(* IEC 61131-3 sources: 2026_Projet_YGO_ExcavatriceDragage/TOOLS/TEST_AUTO_CI/RESULTS/I_TRANSLATION/reports (part 3) *)

    ASSERT_FALSE(RestartSeen, 'aucun front montant mot/frequence apres l armement du verrou');
    ASSERT_TRUE(FB_T.ArrivalStopConfirmed, 'l arret confirme resiste au rebond et a la re-demande');
END_TEST

TEST 'TC-P11-037 T345-L1 Le fait d arret confirme n est ni constant ni efface par la demande'
    CfgFast.CfgRampAccelRate := 1000.0;
    CfgFast.CfgRampDecelNormalRate := 1000.0;
    CfgFast.CaptorDebounce := T#100ms;
    CfgFast.BrakeDelayMagnetise := T#0ms;
    CfgFast.BrakeDelayContactClose := T#0ms;

    (* Scan 1 : au repos, aucun arret confirme (le fait n est pas constant) *)
    FB_T(Enable := TRUE, Reset := FALSE, RunRequest := FALSE, SafeStop := FALSE,
         ReqTremie := FALSE, ReqMaintenance := FALSE, SpeedTgt_Pct := 50.0,
         PowerContactorEngaged := TRUE, Cfg := CfgFast,
         BypassContactorCheck := TRUE, BrakeFeedback := TRUE);
    ASSERT_FALSE(FB_T.ArrivalStopConfirmed, 'au repos : aucun arret confirme (fait non constant)');
    ADVANCE_TIME(10000000);

    (* Scans 2-5 : mouvement vers la cible *)
    FB_T(Enable := TRUE, Reset := FALSE, RunRequest := TRUE, SafeStop := FALSE,
         ReqTremie := TRUE, ReqMaintenance := FALSE, EffectivePermitM3_Tremie := TRUE,
         SpeedTgt_Pct := 50.0, PowerContactorEngaged := TRUE, Cfg := CfgFast,
         BypassContactorCheck := TRUE, BrakeFeedback := TRUE);
    ADVANCE_TIME(10000000);
    FB_T(Enable := TRUE, Reset := FALSE, RunRequest := TRUE, SafeStop := FALSE,
         ReqTremie := TRUE, ReqMaintenance := FALSE, EffectivePermitM3_Tremie := TRUE,
         SpeedTgt_Pct := 50.0, PowerContactorEngaged := TRUE, Cfg := CfgFast,
         BypassContactorCheck := TRUE, BrakeFeedback := TRUE);
    ADVANCE_TIME(10000000);
    FB_T(Enable := TRUE, Reset := FALSE, RunRequest := TRUE, SafeStop := FALSE,
         ReqTremie := TRUE, ReqMaintenance := FALSE, EffectivePermitM3_Tremie := TRUE,
         SpeedTgt_Pct := 50.0, PowerContactorEngaged := TRUE, Cfg := CfgFast,
         BypassContactorCheck := TRUE, BrakeFeedback := TRUE);
    ADVANCE_TIME(10000000);
    FB_T(Enable := TRUE, Reset := FALSE, RunRequest := TRUE, SafeStop := FALSE,
         ReqTremie := TRUE, ReqMaintenance := FALSE, EffectivePermitM3_Tremie := TRUE,
         SpeedTgt_Pct := 50.0, PowerContactorEngaged := TRUE, Cfg := CfgFast,
         BypassContactorCheck := TRUE, BrakeFeedback := TRUE);
    ASSERT_FALSE(FB_T.ArrivalStopConfirmed, 'en mouvement : aucun arret confirme');
    ADVANCE_TIME(10000000);

    (* Scans 6-20 : capteur cible, puis demande retiree avant la fin du debounce *)
    FB_T(Enable := TRUE, Reset := FALSE, RunRequest := TRUE, SafeStop := FALSE,
         ReqTremie := TRUE, ReqMaintenance := FALSE, EffectivePermitM3_Tremie := TRUE,
         SpeedTgt_Pct := 50.0, PowerContactorEngaged := TRUE, PositionSensorTarget := TRUE,
         Cfg := CfgFast, BypassContactorCheck := TRUE, BrakeFeedback := TRUE);
    ADVANCE_TIME(10000000);
    FB_T(Enable := TRUE, Reset := FALSE, RunRequest := FALSE, SafeStop := FALSE,
         ReqTremie := FALSE, ReqMaintenance := FALSE, EffectivePermitM3_Tremie := TRUE,
         SpeedTgt_Pct := 50.0, PowerContactorEngaged := TRUE, PositionSensorTarget := TRUE,
         Cfg := CfgFast, BypassContactorCheck := TRUE, BrakeFeedback := TRUE);
    ADVANCE_TIME(10000000);
    FB_T(Enable := TRUE, Reset := FALSE, RunRequest := FALSE, SafeStop := FALSE,
         ReqTremie := FALSE, ReqMaintenance := FALSE, EffectivePermitM3_Tremie := TRUE,
         SpeedTgt_Pct := 50.0, PowerContactorEngaged := TRUE, PositionSensorTarget := TRUE,
         Cfg := CfgFast, BypassContactorCheck := TRUE, BrakeFeedback := TRUE);
    ADVANCE_TIME(10000000);
    FB_T(Enable := TRUE, Reset := FALSE, RunRequest := FALSE, SafeStop := FALSE,
         ReqTremie := FALSE, ReqMaintenance := FALSE, EffectivePermitM3_Tremie := TRUE,
         SpeedTgt_Pct := 50.0, PowerContactorEngaged := TRUE, PositionSensorTarget := TRUE,
         Cfg := CfgFast, BypassContactorCheck := TRUE, BrakeFeedback := TRUE);
    ADVANCE_TIME(10000000);
    FB_T(Enable := TRUE, Reset := FALSE, RunRequest := FALSE, SafeStop := FALSE,
         ReqTremie := FALSE, ReqMaintenance := FALSE, EffectivePermitM3_Tremie := TRUE,
         SpeedTgt_Pct := 50.0, PowerContactorEngaged := TRUE, PositionSensorTarget := TRUE,
         Cfg := CfgFast, BypassContactorCheck := TRUE, BrakeFeedback := TRUE);
    ADVANCE_TIME(10000000);
    FB_T(Enable := TRUE, Reset := FALSE, RunRequest := FALSE, SafeStop := FALSE,
         ReqTremie := FALSE, ReqMaintenance := FALSE, EffectivePermitM3_Tremie := TRUE,
         SpeedTgt_Pct := 50.0, PowerContactorEngaged := TRUE, PositionSensorTarget := TRUE,
         Cfg := CfgFast, BypassContactorCheck := TRUE, BrakeFeedback := TRUE);
    ADVANCE_TIME(10000000);
    FB_T(Enable := TRUE, Reset := FALSE, RunRequest := FALSE, SafeStop := FALSE,
         ReqTremie := FALSE, ReqMaintenance := FALSE, EffectivePermitM3_Tremie := TRUE,
         SpeedTgt_Pct := 50.0, PowerContactorEngaged := TRUE, PositionSensorTarget := TRUE,
         Cfg := CfgFast, BypassContactorCheck := TRUE, BrakeFeedback := TRUE);
    ADVANCE_TIME(10000000);
    FB_T(Enable := TRUE, Reset := FALSE, RunRequest := FALSE, SafeStop := FALSE,
         ReqTremie := FALSE, ReqMaintenance := FALSE, EffectivePermitM3_Tremie := TRUE,
         SpeedTgt_Pct := 50.0, PowerContactorEngaged := TRUE, PositionSensorTarget := TRUE,
         Cfg := CfgFast, BypassContactorCheck := TRUE, BrakeFeedback := TRUE);
    ADVANCE_TIME(10000000);
    FB_T(Enable := TRUE, Reset := FALSE, RunRequest := FALSE, SafeStop := FALSE,
         ReqTremie := FALSE, ReqMaintenance := FALSE, EffectivePermitM3_Tremie := TRUE,
         SpeedTgt_Pct := 50.0, PowerContactorEngaged := TRUE, PositionSensorTarget := TRUE,
         Cfg := CfgFast, BypassContactorCheck := TRUE, BrakeFeedback := TRUE);
    ADVANCE_TIME(10000000);
    FB_T(Enable := TRUE, Reset := FALSE, RunRequest := FALSE, SafeStop := FALSE,
         ReqTremie := FALSE, ReqMaintenance := FALSE, EffectivePermitM3_Tremie := TRUE,
         SpeedTgt_Pct := 50.0, PowerContactorEngaged := TRUE, PositionSensorTarget := TRUE,
         Cfg := CfgFast, BypassContactorCheck := TRUE, BrakeFeedback := TRUE);
    ADVANCE_TIME(10000000);
    FB_T(Enable := TRUE, Reset := FALSE, RunRequest := FALSE, SafeStop := FALSE,
         ReqTremie := FALSE, ReqMaintenance := FALSE, EffectivePermitM3_Tremie := TRUE,
         SpeedTgt_Pct := 50.0, PowerContactorEngaged := TRUE, PositionSensorTarget := TRUE,
         Cfg := CfgFast, BypassContactorCheck := TRUE, BrakeFeedback := TRUE);
    ADVANCE_TIME(10000000);
    FB_T(Enable := TRUE, Reset := FALSE, RunRequest := FALSE, SafeStop := FALSE,
         ReqTremie := FALSE, ReqMaintenance := FALSE, EffectivePermitM3_Tremie := TRUE,
         SpeedTgt_Pct := 50.0, PowerContactorEngaged := TRUE, PositionSensorTarget := TRUE,
         Cfg := CfgFast, BypassContactorCheck := TRUE, BrakeFeedback := TRUE);
    ADVANCE_TIME(10000000);
    FB_T(Enable := TRUE, Reset := FALSE, RunRequest := FALSE, SafeStop := FALSE,
         ReqTremie := FALSE, ReqMaintenance := FALSE, EffectivePermitM3_Tremie := TRUE,
         SpeedTgt_Pct := 50.0, PowerContactorEngaged := TRUE, PositionSensorTarget := TRUE,
         Cfg := CfgFast, BypassContactorCheck := TRUE, BrakeFeedback := TRUE);
    ADVANCE_TIME(10000000);
    FB_T(Enable := TRUE, Reset := FALSE, RunRequest := FALSE, SafeStop := FALSE,
         ReqTremie := FALSE, ReqMaintenance := FALSE, EffectivePermitM3_Tremie := TRUE,
         SpeedTgt_Pct := 50.0, PowerContactorEngaged := TRUE, PositionSensorTarget := TRUE,
         Cfg := CfgFast, BypassContactorCheck := TRUE, BrakeFeedback := TRUE);
    ADVANCE_TIME(10000000);
    FB_T(Enable := TRUE, Reset := FALSE, RunRequest := FALSE, SafeStop := FALSE,
         ReqTremie := FALSE, ReqMaintenance := FALSE, EffectivePermitM3_Tremie := TRUE,
         SpeedTgt_Pct := 50.0, PowerContactorEngaged := TRUE, PositionSensorTarget := TRUE,
         Cfg := CfgFast, BypassContactorCheck := TRUE, BrakeFeedback := TRUE);
    ADVANCE_TIME(10000000);
    ASSERT_TRUE(FB_T.ArrivalStopConfirmed, 'demande retiree avant le debounce : arret confirme');

    (* Scans 21-24 : la demande du MEME sens est re-armee, cible stable -> le fait doit tenir *)
    FB_T(Enable := TRUE, Reset := FALSE, RunRequest := TRUE, SafeStop := FALSE,
         ReqTremie := TRUE, ReqMaintenance := FALSE, EffectivePermitM3_Tremie := TRUE,
         SpeedTgt_Pct := 50.0, PowerContactorEngaged := TRUE, PositionSensorTarget := TRUE,
         Cfg := CfgFast, BypassContactorCheck := TRUE, BrakeFeedback := TRUE);
    ADVANCE_TIME(10000000);
    FB_T(Enable := TRUE, Reset := FALSE, RunRequest := TRUE, SafeStop := FALSE,
         ReqTremie := TRUE, ReqMaintenance := FALSE, EffectivePermitM3_Tremie := TRUE,
         SpeedTgt_Pct := 50.0, PowerContactorEngaged := TRUE, PositionSensorTarget := TRUE,
         Cfg := CfgFast, BypassContactorCheck := TRUE, BrakeFeedback := TRUE);
    ADVANCE_TIME(10000000);
    FB_T(Enable := TRUE, Reset := FALSE, RunRequest := TRUE, SafeStop := FALSE,
         ReqTremie := TRUE, ReqMaintenance := FALSE, EffectivePermitM3_Tremie := TRUE,
         SpeedTgt_Pct := 50.0, PowerContactorEngaged := TRUE, PositionSensorTarget := TRUE,
         Cfg := CfgFast, BypassContactorCheck := TRUE, BrakeFeedback := TRUE);
    ADVANCE_TIME(10000000);
    FB_T(Enable := TRUE, Reset := FALSE, RunRequest := TRUE, SafeStop := FALSE,
         ReqTremie := TRUE, ReqMaintenance := FALSE, EffectivePermitM3_Tremie := TRUE,
         SpeedTgt_Pct := 50.0, PowerContactorEngaged := TRUE, PositionSensorTarget := TRUE,
         Cfg := CfgFast, BypassContactorCheck := TRUE, BrakeFeedback := TRUE);
    ASSERT_TRUE(FB_T.ArrivalStopConfirmed, 're-demande du meme sens : arret confirme conserve');
    ASSERT_EQ(FB_T.RequestedDriveControlWord, 0, 're-demande du meme sens : mot de commande reste a 0');
END_TEST

TEST 'TC-P11-038 T345-L1 Une demande de SENS INVERSE relache le verrou et autorise le degagement'
    CfgFast.CfgRampAccelRate := 1000.0;
    CfgFast.CfgRampDecelNormalRate := 1000.0;
    CfgFast.BrakeDelayMagnetise := T#0ms;
    CfgFast.BrakeDelayContactClose := T#0ms;

    (* Scans 1-4 : mouvement vers la cible puis capteur cible + demande retiree *)
    FB_T(Enable := TRUE, Reset := FALSE, RunRequest := TRUE, SafeStop := FALSE,
         ReqTremie := TRUE, ReqMaintenance := FALSE, EffectivePermitM3_Tremie := TRUE,
         SpeedTgt_Pct := 50.0, PowerContactorEngaged := TRUE, Cfg := CfgFast,
         BypassContactorCheck := TRUE, BrakeFeedback := TRUE);
    ADVANCE_TIME(10000000);
    FB_T(Enable := TRUE, Reset := FALSE, RunRequest := TRUE, SafeStop := FALSE,
         ReqTremie := TRUE, ReqMaintenance := FALSE, EffectivePermitM3_Tremie := TRUE,
         SpeedTgt_Pct := 50.0, PowerContactorEngaged := TRUE, Cfg := CfgFast,
         BypassContactorCheck := TRUE, BrakeFeedback := TRUE);
    ADVANCE_TIME(10000000);
    FB_T(Enable := TRUE, Reset := FALSE, RunRequest := TRUE, SafeStop := FALSE,
         ReqTremie := TRUE, ReqMaintenance := FALSE, EffectivePermitM3_Tremie := TRUE,
         SpeedTgt_Pct := 50.0, PowerContactorEngaged := TRUE, Cfg := CfgFast,
         BypassContactorCheck := TRUE, BrakeFeedback := TRUE);
    ADVANCE_TIME(10000000);
    FB_T(Enable := TRUE, Reset := FALSE, RunRequest := TRUE, SafeStop := FALSE,
         ReqTremie := TRUE, ReqMaintenance := FALSE, EffectivePermitM3_Tremie := TRUE,
         SpeedTgt_Pct := 50.0, PowerContactorEngaged := TRUE, PositionSensorTarget := TRUE,
         Cfg := CfgFast, BypassContactorCheck := TRUE, BrakeFeedback := TRUE);
    ADVANCE_TIME(10000000);
    FB_T(Enable := TRUE, Reset := FALSE, RunRequest := FALSE, SafeStop := FALSE,
         ReqTremie := FALSE, ReqMaintenance := FALSE, EffectivePermitM3_Tremie := TRUE,
         SpeedTgt_Pct := 50.0, PowerContactorEngaged := TRUE, PositionSensorTarget := TRUE,
         Cfg := CfgFast, BypassContactorCheck := TRUE, BrakeFeedback := TRUE);
    ADVANCE_TIME(10000000);
    FB_T(Enable := TRUE, Reset := FALSE, RunRequest := FALSE, SafeStop := FALSE,
         ReqTremie := FALSE, ReqMaintenance := FALSE, EffectivePermitM3_Tremie := TRUE,
         SpeedTgt_Pct := 50.0, PowerContactorEngaged := TRUE, PositionSensorTarget := TRUE,
         Cfg := CfgFast, BypassContactorCheck := TRUE, BrakeFeedback := TRUE);
    ADVANCE_TIME(10000000);
    FB_T(Enable := TRUE, Reset := FALSE, RunRequest := FALSE, SafeStop := FALSE,
         ReqTremie := FALSE, ReqMaintenance := FALSE, EffectivePermitM3_Tremie := TRUE,
         SpeedTgt_Pct := 50.0, PowerContactorEngaged := TRUE, PositionSensorTarget := TRUE,
         Cfg := CfgFast, BypassContactorCheck := TRUE, BrakeFeedback := TRUE);
    ADVANCE_TIME(10000000);
    FB_T(Enable := TRUE, Reset := FALSE, RunRequest := FALSE, SafeStop := FALSE,
         ReqTremie := FALSE, ReqMaintenance := FALSE, EffectivePermitM3_Tremie := TRUE,
         SpeedTgt_Pct := 50.0, PowerContactorEngaged := TRUE, PositionSensorTarget := TRUE,
         Cfg := CfgFast, BypassContactorCheck := TRUE, BrakeFeedback := TRUE);
    ADVANCE_TIME(10000000);
    FB_T(Enable := TRUE, Reset := FALSE, RunRequest := FALSE, SafeStop := FALSE,
         ReqTremie := FALSE, ReqMaintenance := FALSE, EffectivePermitM3_Tremie := TRUE,
         SpeedTgt_Pct := 50.0, PowerContactorEngaged := TRUE, PositionSensorTarget := TRUE,
         Cfg := CfgFast, BypassContactorCheck := TRUE, BrakeFeedback := TRUE);
    ADVANCE_TIME(10000000);
    FB_T(Enable := TRUE, Reset := FALSE, RunRequest := FALSE, SafeStop := FALSE,
         ReqTremie := FALSE, ReqMaintenance := FALSE, EffectivePermitM3_Tremie := TRUE,
         SpeedTgt_Pct := 50.0, PowerContactorEngaged := TRUE, PositionSensorTarget := TRUE,
         Cfg := CfgFast, BypassContactorCheck := TRUE, BrakeFeedback := TRUE);
    ADVANCE_TIME(10000000);
    FB_T(Enable := TRUE, Reset := FALSE, RunRequest := FALSE, SafeStop := FALSE,
         ReqTremie := FALSE, ReqMaintenance := FALSE, EffectivePermitM3_Tremie := TRUE,
         SpeedTgt_Pct := 50.0, PowerContactorEngaged := TRUE, PositionSensorTarget := TRUE,
         Cfg := CfgFast, BypassContactorCheck := TRUE, BrakeFeedback := TRUE);
    ADVANCE_TIME(10000000);
    FB_T(Enable := TRUE, Reset := FALSE, RunRequest := FALSE, SafeStop := FALSE,
         ReqTremie := FALSE, ReqMaintenance := FALSE, EffectivePermitM3_Tremie := TRUE,
         SpeedTgt_Pct := 50.0, PowerContactorEngaged := TRUE, PositionSensorTarget := TRUE,
         Cfg := CfgFast, BypassContactorCheck := TRUE, BrakeFeedback := TRUE);
    ADVANCE_TIME(10000000);
    FB_T(Enable := TRUE, Reset := FALSE, RunRequest := FALSE, SafeStop := FALSE,
         ReqTremie := FALSE, ReqMaintenance := FALSE, EffectivePermitM3_Tremie := TRUE,
         SpeedTgt_Pct := 50.0, PowerContactorEngaged := TRUE, PositionSensorTarget := TRUE,
         Cfg := CfgFast, BypassContactorCheck := TRUE, BrakeFeedback := TRUE);
    ADVANCE_TIME(10000000);
    FB_T(Enable := TRUE, Reset := FALSE, RunRequest := FALSE, SafeStop := FALSE,
         ReqTremie := FALSE, ReqMaintenance := FALSE, EffectivePermitM3_Tremie := TRUE,
         SpeedTgt_Pct := 50.0, PowerContactorEngaged := TRUE, PositionSensorTarget := TRUE,
         Cfg := CfgFast, BypassContactorCheck := TRUE, BrakeFeedback := TRUE);
    ASSERT_TRUE(FB_T.ArrivalStopConfirmed, 'verrou d arret arme avec le sens du mouvement');
    ADVANCE_TIME(10000000);

    (* Scans 15-18 : demande explicite de SENS INVERSE (Maintenance) -> degagement autorise *)
    FB_T(Enable := TRUE, Reset := FALSE, RunRequest := TRUE, SafeStop := FALSE,
         ReqTremie := FALSE, ReqMaintenance := TRUE, EffectivePermitM3_Maintenance := TRUE,
         SpeedTgt_Pct := 50.0, PowerContactorEngaged := TRUE, PositionSensorTarget := TRUE,
         Cfg := CfgFast, BypassContactorCheck := TRUE, BrakeFeedback := TRUE);
    ADVANCE_TIME(10000000);
    FB_T(Enable := TRUE, Reset := FALSE, RunRequest := TRUE, SafeStop := FALSE,
         ReqTremie := FALSE, ReqMaintenance := TRUE, EffectivePermitM3_Maintenance := TRUE,
         SpeedTgt_Pct := 50.0, PowerContactorEngaged := TRUE, PositionSensorTarget := TRUE,
         Cfg := CfgFast, BypassContactorCheck := TRUE, BrakeFeedback := TRUE);
    ADVANCE_TIME(10000000);
    FB_T(Enable := TRUE, Reset := FALSE, RunRequest := TRUE, SafeStop := FALSE,
         ReqTremie := FALSE, ReqMaintenance := TRUE, EffectivePermitM3_Maintenance := TRUE,
         SpeedTgt_Pct := 50.0, PowerContactorEngaged := TRUE, PositionSensorTarget := TRUE,
         Cfg := CfgFast, BypassContactorCheck := TRUE, BrakeFeedback := TRUE);
    ADVANCE_TIME(10000000);
    FB_T(Enable := TRUE, Reset := FALSE, RunRequest := TRUE, SafeStop := FALSE,
         ReqTremie := FALSE, ReqMaintenance := TRUE, EffectivePermitM3_Maintenance := TRUE,
         SpeedTgt_Pct := 50.0, PowerContactorEngaged := TRUE, PositionSensorTarget := TRUE,
         Cfg := CfgFast, BypassContactorCheck := TRUE, BrakeFeedback := TRUE);
    ASSERT_EQ(FB_T.RequestedDriveControlWord, 2, 'sens inverse : mot de commande REV');
    ASSERT_GT(FB_T.RequestedDriveFreqHz, 0.0, 'sens inverse : consigne de frequence non nulle');
    ASSERT_FALSE(FB_T.ArrivalStopConfirmed, 'axe en mouvement : plus d arret confirme');
END_TEST

TEST 'TC-P11-039 T345-L1 Non-vacuite : rotation reelle au variateur -> aucun arret confirme'
    CfgFast.CfgRampAccelRate := 1000.0;
    CfgFast.CfgRampDecelNormalRate := 1000.0;
    CfgFast.BrakeDelayMagnetise := T#0ms;
    CfgFast.BrakeDelayContactClose := T#0ms;

    (* Scans 1-4 : mouvement vers la cible *)
    FB_T(Enable := TRUE, Reset := FALSE, RunRequest := TRUE, SafeStop := FALSE,
         ReqTremie := TRUE, ReqMaintenance := FALSE, EffectivePermitM3_Tremie := TRUE,
         SpeedTgt_Pct := 50.0, PowerContactorEngaged := TRUE, Cfg := CfgFast,
         BypassContactorCheck := TRUE, BrakeFeedback := TRUE);
    ADVANCE_TIME(10000000);
    FB_T(Enable := TRUE, Reset := FALSE, RunRequest := TRUE, SafeStop := FALSE,
         ReqTremie := TRUE, ReqMaintenance := FALSE, EffectivePermitM3_Tremie := TRUE,
         SpeedTgt_Pct := 50.0, PowerContactorEngaged := TRUE, Cfg := CfgFast,
         BypassContactorCheck := TRUE, BrakeFeedback := TRUE);
    ADVANCE_TIME(10000000);
    FB_T(Enable := TRUE, Reset := FALSE, RunRequest := TRUE, SafeStop := FALSE,
         ReqTremie := TRUE, ReqMaintenance := FALSE, EffectivePermitM3_Tremie := TRUE,
         SpeedTgt_Pct := 50.0, PowerContactorEngaged := TRUE, Cfg := CfgFast,
         BypassContactorCheck := TRUE, BrakeFeedback := TRUE);
    ADVANCE_TIME(10000000);
    FB_T(Enable := TRUE, Reset := FALSE, RunRequest := TRUE, SafeStop := FALSE,
         ReqTremie := TRUE, ReqMaintenance := FALSE, EffectivePermitM3_Tremie := TRUE,
         SpeedTgt_Pct := 50.0, PowerContactorEngaged := TRUE, PositionSensorTarget := TRUE,
         Cfg := CfgFast, BypassContactorCheck := TRUE, BrakeFeedback := TRUE);
    ADVANCE_TIME(10000000);

    (* Scans 5-18 : demande retiree, cible tenue -> arret confirme *)
    FB_T(Enable := TRUE, Reset := FALSE, RunRequest := FALSE, SafeStop := FALSE,
         ReqTremie := FALSE, ReqMaintenance := FALSE, SpeedTgt_Pct := 50.0,
         PowerContactorEngaged := TRUE, PositionSensorTarget := TRUE,
         Cfg := CfgFast, BypassContactorCheck := TRUE, BrakeFeedback := TRUE);
    ADVANCE_TIME(10000000);
    FB_T(Enable := TRUE, Reset := FALSE, RunRequest := FALSE, SafeStop := FALSE,
         ReqTremie := FALSE, ReqMaintenance := FALSE, SpeedTgt_Pct := 50.0,
         PowerContactorEngaged := TRUE, PositionSensorTarget := TRUE,
         Cfg := CfgFast, BypassContactorCheck := TRUE, BrakeFeedback := TRUE);
    ADVANCE_TIME(10000000);
    FB_T(Enable := TRUE, Reset := FALSE, RunRequest := FALSE, SafeStop := FALSE,
         ReqTremie := FALSE, ReqMaintenance := FALSE, SpeedTgt_Pct := 50.0,
         PowerContactorEngaged := TRUE, PositionSensorTarget := TRUE,
         Cfg := CfgFast, BypassContactorCheck := TRUE, BrakeFeedback := TRUE);
    ADVANCE_TIME(10000000);
    FB_T(Enable := TRUE, Reset := FALSE, RunRequest := FALSE, SafeStop := FALSE,
         ReqTremie := FALSE, ReqMaintenance := FALSE, SpeedTgt_Pct := 50.0,
         PowerContactorEngaged := TRUE, PositionSensorTarget := TRUE,
         Cfg := CfgFast, BypassContactorCheck := TRUE, BrakeFeedback := TRUE);
    ADVANCE_TIME(10000000);
    FB_T(Enable := TRUE, Reset := FALSE, RunRequest := FALSE, SafeStop := FALSE,
         ReqTremie := FALSE, ReqMaintenance := FALSE, SpeedTgt_Pct := 50.0,
         PowerContactorEngaged := TRUE, PositionSensorTarget := TRUE,
         Cfg := CfgFast, BypassContactorCheck := TRUE, BrakeFeedback := TRUE);
    ADVANCE_TIME(10000000);
    FB_T(Enable := TRUE, Reset := FALSE, RunRequest := FALSE, SafeStop := FALSE,
         ReqTremie := FALSE, ReqMaintenance := FALSE, SpeedTgt_Pct := 50.0,
         PowerContactorEngaged := TRUE, PositionSensorTarget := TRUE,
         Cfg := CfgFast, BypassContactorCheck := TRUE, BrakeFeedback := TRUE);
    ADVANCE_TIME(10000000);
    FB_T(Enable := TRUE, Reset := FALSE, RunRequest := FALSE, SafeStop := FALSE,
         ReqTremie := FALSE, ReqMaintenance := FALSE, SpeedTgt_Pct := 50.0,
         PowerContactorEngaged := TRUE, PositionSensorTarget := TRUE,
         Cfg := CfgFast, BypassContactorCheck := TRUE, BrakeFeedback := TRUE);
    ADVANCE_TIME(10000000);
    FB_T(Enable := TRUE, Reset := FALSE, RunRequest := FALSE, SafeStop := FALSE,
         ReqTremie := FALSE, ReqMaintenance := FALSE, SpeedTgt_Pct := 50.0,
         PowerContactorEngaged := TRUE, PositionSensorTarget := TRUE,
         Cfg := CfgFast, BypassContactorCheck := TRUE, BrakeFeedback := TRUE);
    ADVANCE_TIME(10000000);
    FB_T(Enable := TRUE, Reset := FALSE, RunRequest := FALSE, SafeStop := FALSE,
         ReqTremie := FALSE, ReqMaintenance := FALSE, SpeedTgt_Pct := 50.0,
         PowerContactorEngaged := TRUE, PositionSensorTarget := TRUE,
         Cfg := CfgFast, BypassContactorCheck := TRUE, BrakeFeedback := TRUE);
    ADVANCE_TIME(10000000);
    FB_T(Enable := TRUE, Reset := FALSE, RunRequest := FALSE, SafeStop := FALSE,
         ReqTremie := FALSE, ReqMaintenance := FALSE, SpeedTgt_Pct := 50.0,
         PowerContactorEngaged := TRUE, PositionSensorTarget := TRUE,
         Cfg := CfgFast, BypassContactorCheck := TRUE, BrakeFeedback := TRUE);
    ADVANCE_TIME(10000000);
    FB_T(Enable := TRUE, Reset := FALSE, RunRequest := FALSE, SafeStop := FALSE,
         ReqTremie := FALSE, ReqMaintenance := FALSE, SpeedTgt_Pct := 50.0,
         PowerContactorEngaged := TRUE, PositionSensorTarget := TRUE,
         Cfg := CfgFast, BypassContactorCheck := TRUE, BrakeFeedback := TRUE);
    ADVANCE_TIME(10000000);
    FB_T(Enable := TRUE, Reset := FALSE, RunRequest := FALSE, SafeStop := FALSE,
         ReqTremie := FALSE, ReqMaintenance := FALSE, SpeedTgt_Pct := 50.0,
         PowerContactorEngaged := TRUE, PositionSensorTarget := TRUE,
         Cfg := CfgFast, BypassContactorCheck := TRUE, BrakeFeedback := TRUE);
    ADVANCE_TIME(10000000);
    FB_T(Enable := TRUE, Reset := FALSE, RunRequest := FALSE, SafeStop := FALSE,
         ReqTremie := FALSE, ReqMaintenance := FALSE, SpeedTgt_Pct := 50.0,
         PowerContactorEngaged := TRUE, PositionSensorTarget := TRUE,
         Cfg := CfgFast, BypassContactorCheck := TRUE, BrakeFeedback := TRUE);
    ADVANCE_TIME(10000000);
    FB_T(Enable := TRUE, Reset := FALSE, RunRequest := FALSE, SafeStop := FALSE,
         ReqTremie := FALSE, ReqMaintenance := FALSE, SpeedTgt_Pct := 50.0,
         PowerContactorEngaged := TRUE, PositionSensorTarget := TRUE, DriveActualFreqHz := 0.0,
         Cfg := CfgFast, BypassContactorCheck := TRUE, BrakeFeedback := TRUE);
    ASSERT_TRUE(FB_T.ArrivalStopConfirmed, 'arret au repos : fait publie');
    ADVANCE_TIME(10000000);

    (* Scan 19 : le variateur tourne encore (5,0 Hz) -> l arret n est PAS confirme *)
    FB_T(Enable := TRUE, Reset := FALSE, RunRequest := FALSE, SafeStop := FALSE,
         ReqTremie := FALSE, ReqMaintenance := FALSE, SpeedTgt_Pct := 50.0,
         PowerContactorEngaged := TRUE, PositionSensorTarget := TRUE, DriveActualFreqHz := 5.0,
         Cfg := CfgFast, BypassContactorCheck := TRUE, BrakeFeedback := TRUE);
    ASSERT_FALSE(FB_T.ArrivalStopConfirmed, 'rotation reelle 5,0 Hz : aucun arret confirme');
    ADVANCE_TIME(10000000);

    (* Scan 20 : retour au repos reel -> fait de nouveau publie *)
    FB_T(Enable := TRUE, Reset := FALSE, RunRequest := FALSE, SafeStop := FALSE,
         ReqTremie := FALSE, ReqMaintenance := FALSE, SpeedTgt_Pct := 50.0,
         PowerContactorEngaged := TRUE, PositionSensorTarget := TRUE, DriveActualFreqHz := 0.0,
         Cfg := CfgFast, BypassContactorCheck := TRUE, BrakeFeedback := TRUE);
    ASSERT_TRUE(FB_T.ArrivalStopConfirmed, 'retour au repos : arret confirme publie');
END_TEST

(* ---- FB_TranslationOutputInterlock_test.st ---- *)
(* =======================================================================
   Automated Unit Test - FB_TranslationOutputInterlock
   ======================================================================= *)
TEST 'TC-P11-INT-001 Enable FALSE coupe consignes variateur et ordre frein'
VAR
    fb : FB_TranslationOutputInterlock;
END_VAR
    fb.Enable := FALSE;
    fb.RequestedDriveControlWord := 1; (* Fwd *)
    fb.RequestedDriveFreqHz := 50.0;
    fb.BrakeReleaseRequest := TRUE;
    fb();
    ASSERT_FALSE(fb.Ready, 'Enable FALSE -> Ready FALSE');
    ASSERT_EQ(fb.DriveControlWord, 0, 'Enable FALSE -> Mot variateur 0');
    ASSERT_EQ(fb.DriveFreqCmd_Hz, 0.0, 'Enable FALSE -> Frequence 0.0');
    ASSERT_FALSE(fb.BrakeCmd, 'Enable FALSE -> Frein non desserre');
END_TEST

TEST 'TC-P11-INT-002 Blocage sens sans permis directionnel (fail-safe)'
VAR
    fb : FB_TranslationOutputInterlock;
END_VAR
    fb.Enable := TRUE;
    fb.PowerContactorEngaged := TRUE;
    fb.EffectivePermitM3_Tremie := FALSE; (* Permis Tremie refuse *)
    fb.RequestedDriveControlWord := 1; (* Demande Fwd Tremie *)
    fb.RequestedDriveFreqHz := 25.0;
    fb();
    ASSERT_EQ(fb.DriveControlWord, 0, 'Permis Tremie FALSE -> Mot bloque a 0');
    ASSERT_EQ(fb.DriveFreqCmd_Hz, 0.0, 'Permis Tremie FALSE -> Frequence bloquee a 0.0');
END_TEST

TEST 'TC-P11-INT-003 Mouvement nominal autorise avec permis et confirmation frein'
VAR
    fb : FB_TranslationOutputInterlock;
END_VAR
    fb.Enable := TRUE;
    fb.PowerContactorEngaged := TRUE;
    fb.EffectivePermitM3_Tremie := TRUE;
    fb.BrakeReleaseRequest := TRUE;
    fb.BrakeCommandOpenConfirmed := TRUE; (* Frein ouvert confirme *)
    fb.RequestedDriveControlWord := 1; (* Fwd Tremie *)
    fb.RequestedDriveFreqHz := 30.0;
    fb();
    ASSERT_TRUE(fb.Ready, 'Conditions OK -> Ready TRUE');
    ASSERT_EQ(fb.DriveControlWord, 1, 'Permis OK + Frein OK -> Mot Fwd emis');
    ASSERT_EQ(fb.DriveFreqCmd_Hz, 30.0, 'Permis OK + Frein OK -> Frequence 30.0');
    ASSERT_TRUE(fb.BrakeCmd, 'BrakeReleaseRequest -> BrakeCmd TRUE');
END_TEST
